// TIA Portal V20 export
// export: Created 2026-10-20T12:44:49.8654744Z, ExportSetting WithDefaults, DisplayName Totally Integrated Automation Portal, DisplayVersion V20 Update 6, DisplayName TIA Portal Openness, DisplayVersion V20 Update 6, DisplayName TIA Portal Version Control Interface, DisplayVersion V20 Update 6, DisplayName SINAMICS Startdrive Advanced, DisplayVersion V20 SP1, DisplayName SINAMICS Startdrive G130, G150, S120, S150, SINAMICS MV, G220, S200, S210, DisplayVersion V20 SP1, DisplayName SINAMICS Startdrive G110M, G120, G120C, G120D, G120P, G115D, DisplayVersion V20 SP1, DisplayName STEP 7 Professional, DisplayVersion V20 Update 6, DisplayName STEP 7 Safety, DisplayVersion V20 Update 2, DisplayName WinCC Basic/Comfort/Advanced, DisplayVersion V20 Update 6, DisplayName WinCC Unified, DisplayVersion V20 Update 6
FUNCTION "VTD_Charge_Settings" : Void   // FC41, SCL
{ S7_Optimized_Access := 'TRUE' }
VERSION : 0.1
// stored: AutoNumber true, IsIECCheckEnabled false, SetENOAutomatically false, UDAEnableTagReadback false
BEGIN
   //VTD SETTINGS
   CASE "VTD_System_Selected_HMI" OF
       1:
           "PopUps_DB".VTD_Settings := "Settings_DB".VTD_Sys[1];
       2:
           "PopUps_DB".VTD_Settings := "Settings_DB".VTD_Sys[2];
       3:
           "PopUps_DB".VTD_Settings := "Settings_DB".VTD_Sys[3];
       4:
           "PopUps_DB".VTD_Settings := "Settings_DB".VTD_Sys[4];
       5:
           "PopUps_DB".VTD_Settings := "Settings_DB".VTD_Sys[5];
   END_CASE;
END_FUNCTION
